(* PLC project Vn_int_to_real, Beckhoff Automation GmbH TwinCAT PLC Control 3.5.13.21 *)
(* stored: creationDateTime 1970-01-01T00:00:00 *)

PROGRAM Vn_int_to_real

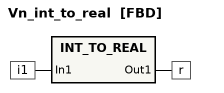
(* FBD diagram, written out as Structured Text *)
r := INT_TO_REAL(i1);
END_PROGRAM
